Fanuc KAREL source: KX00008.KL

PROGRAM KX00008
%NOLOCKGROUP
VAR
  I: INTEGER
  J: INTEGER
  B: BOOLEAN
  F: FILE
  S: STRING[80]
  P: XYZWPR
BEGIN
  ABORT
END KX00008
